SUBAPPLICATION AR_TO_Publish_OPC (* Physikalischer AR-Wert per OPC-UA publiziert, gedrosselt (ohne VT) *)
  (* Standard: 61499-2; Description: Copyright (c) 2026 Meisterschulen am Ostbahnhof This program and the accompanying materials are made available under the terms of the Eclipse Public License 2.0 which is available at https://www.eclipse.org/legal/epl-2.0/ SPDX-License-Identifier: EPL-2.0 *)
  (* Version 1.0, 2026-10-28, Franz Höpfinger, Meisterschulen am Ostbahnhof, Kopie von MyLib::sys::AR_TO_Q_Publish_OPC ohne Q_NumericValue/AR_SPLIT_2, fuer Stationen ohne VT (keine isobus_UT-Libs). RateLimit_Anzeige (500ms) bleibt. *)
  PACKAGE MyLib::sys;
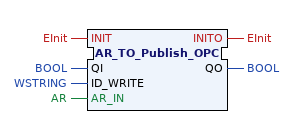
  EVENT_INPUT
    INIT : EInit; (* Initialization Request *)
  END_EVENT
  EVENT_OUTPUT
    INITO : EInit; (* Initialization Confirm *)
  END_EVENT
  VAR_INPUT
    QI : BOOL := TRUE; (* Quality Input - TRUE to enable service *)
    ID_WRITE : WSTRING; (* Publish-Adresse (REAL, ACTION=PUBLISH) *)
  END_VAR
  VAR_OUTPUT
    QO : BOOL; (* Quality Output - TRUE if service executed successfully *)
  END_VAR
  SOCKETS
    AR_IN : adapter::types::unidirectional::AR; (* Physikalischer Wert (bereits skaliert) *)
  END_SOCKETS
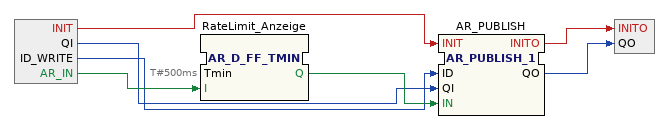
  FBS
    RateLimit_Anzeige : adapter::events::unidirectional::AR_D_FF_TMIN(Tmin := T#500ms); (* Drosselt den Publish auf max. 1 Update/500ms *)
    AR_PUBLISH : adapter::net::AR_PUBLISH_1;
  END_FBS
  EVENT_CONNECTIONS
    INIT TO AR_PUBLISH.INIT;
    AR_PUBLISH.INITO TO INITO;
  END_CONNECTIONS
  DATA_CONNECTIONS
    ID_WRITE TO AR_PUBLISH.ID;
    QI TO AR_PUBLISH.QI;
    AR_PUBLISH.QO TO QO;
  END_CONNECTIONS
  ADAPTER_CONNECTIONS
    AR_IN TO RateLimit_Anzeige.I;
    RateLimit_Anzeige.Q TO AR_PUBLISH.IN;
  END_CONNECTIONS
END_SUBAPPLICATION
